FUNCTION_BLOCK Actuator (* Composite Function Block Type *)
  (* Standard: 61499-2 *)
  (* Version 1.0.1, 10/17/2023, ApplicationLibDevTeam, Schneider Electric, First Version *)
  PACKAGE Flexbridge.FestoMPS400;
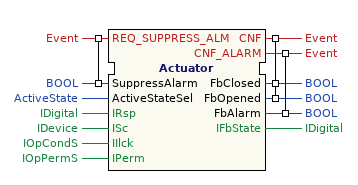
  EVENT_INPUT
    REQ_SUPPRESS_ALM WITH SuppressAlarm; (* Request to update the alarm suppress status *)
  END_EVENT
  EVENT_OUTPUT
    CNF WITH FbClosed, FbOpened; (* Execution confirmation *)
    CNF_ALARM WITH FbAlarm; (* Execution confirmation of alarm *)
  END_EVENT
  VAR_INPUT
    SuppressAlarm : BOOL; (* 1 = Suppress alarm in HMI *)
    ActiveStateSel : ActiveState; (* Feedback type selection to determine the active state for valves [StateSel configured as Valve1Op or Valve2Op],  0 = Open State  1 = Closed State *)
  END_VAR
  VAR_OUTPUT
    FbClosed : BOOL; (* 1 = Closed *)
    FbOpened : BOOL; (* 1 = Opened *)
    FbAlarm : BOOL; (* 1 = Feedback failure alarm is active *)
  END_VAR
  SOCKETS
    IRsp : IDigital; (* Program remote setpoint interface adapter *)
    ISc : IDevice; (* Sequence control Interface adapter. Controls the block when owner is in program local *)
    IIlck : IOpCondS; (* Interlock condition summary chain input from ilckCondItem blocks *)
    IPerm : IOpPermS; (* Permission condition summary chain input from permCondItem blocks *)
  END_SOCKETS
  PLUGS
    IFbState : IDigital; (* Current feedback status adapter(Bit 2 = Feedback failure status) *)
  END_PLUGS
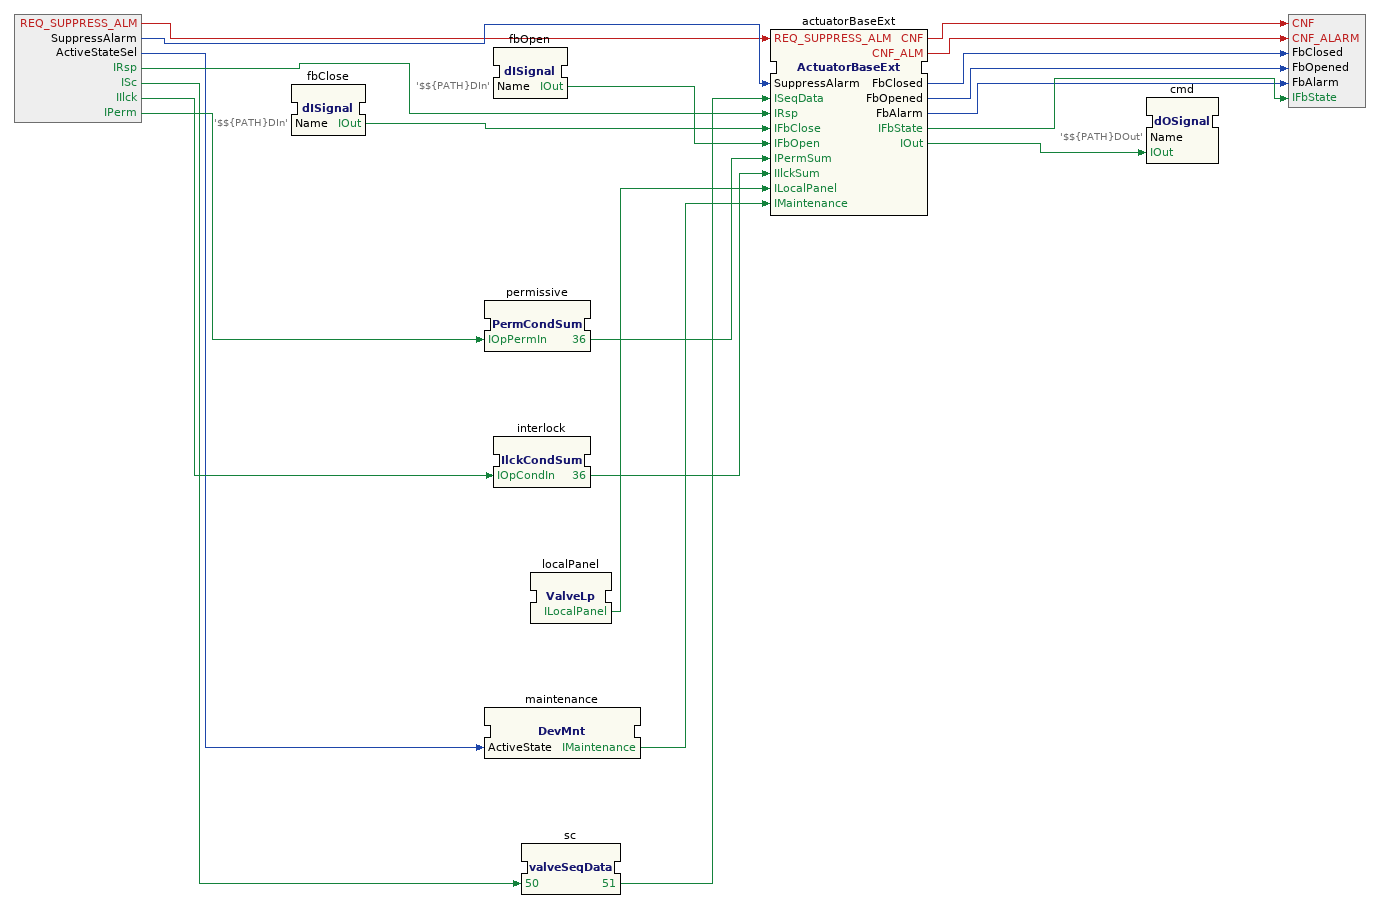
  (* Valve Control *)
  (* Permissive *)
  (* Interlock *)
  (* LocalPanel *)
  (* Maintenance *)
  (* Sequence Control *)
  (* Input Hardware Interface *)
  (* Output Hardware Interface *)
  FBS
    interlock : IlckCondSum; {SET_ATTRIBUTE(Configuration.Component.HideUnusedPorts, )}
    permissive : PermCondSum; {SET_ATTRIBUTE(Configuration.Component.HideUnusedPorts, )}
    localPanel : ValveLp; {SET_ATTRIBUTE(Configuration.Component.HideUnusedPorts, )}
    maintenance : DevMnt; {SET_ATTRIBUTE(Configuration.Component.HideUnusedPorts, )}
    fbOpen : dISignal(Name := '$${PATH}DIn'); {SET_ATTRIBUTE(Configuration.Component.HideUnusedPorts, )}
    cmd : dOSignal(Name := '$${PATH}DOut'); {SET_ATTRIBUTE(Configuration.Component.HideUnusedPorts, )}
    actuatorBaseExt : ActuatorBaseExt;
    fbClose : dISignal(Name := '$${PATH}DIn'); {SET_ATTRIBUTE(Configuration.Component.HideUnusedPorts, )}
    sc : valveSeqData; {SET_ATTRIBUTE(Configuration.Component.HideUnusedPorts, )}
  END_FBS
  EVENT_CONNECTIONS
    actuatorBaseExt.CNF TO CNF;
    actuatorBaseExt.CNF_ALM TO CNF_ALARM;
    REQ_SUPPRESS_ALM TO actuatorBaseExt.REQ_SUPPRESS_ALM;
  END_CONNECTIONS
  DATA_CONNECTIONS
    actuatorBaseExt.FbClosed TO FbClosed;
    actuatorBaseExt.FbOpened TO FbOpened;
    actuatorBaseExt.FbAlarm TO FbAlarm;
    SuppressAlarm TO actuatorBaseExt.SuppressAlarm;
    ActiveStateSel TO maintenance.ActiveState;
  END_CONNECTIONS
  ADAPTER_CONNECTIONS
    IPerm TO permissive.IOpPermIn;
    ISc TO sc.50;
    IIlck TO interlock.IOpCondIn;
    sc.51 TO actuatorBaseExt.ISeqData;
    IRsp TO actuatorBaseExt.IRsp;
    actuatorBaseExt.IFbState TO IFbState;
    actuatorBaseExt.IOut TO cmd.IOut;
    fbClose.IOut TO actuatorBaseExt.IFbClose;
    fbOpen.IOut TO actuatorBaseExt.IFbOpen;
    permissive.36 TO actuatorBaseExt.IPermSum;
    interlock.36 TO actuatorBaseExt.IIlckSum;
    localPanel.ILocalPanel TO actuatorBaseExt.ILocalPanel;
    maintenance.IMaintenance TO actuatorBaseExt.IMaintenance;
  END_CONNECTIONS
END_FUNCTION_BLOCK
